Fanuc KAREL source: kd00051.KL

-- PROVISIONAL review KL for V940-1; original PC SHA256 1b8f119a18a5a4649315fc7f6d6ce60d3f234252100fceed115acb7b17a9f241
-- Incomplete behavior may be omitted. Consult companion uncertainty JSON. Do not deploy.
PROGRAM KD00051
%NOLOCKGROUP
VAR
  I : INTEGER
  J : INTEGER
  B : BOOLEAN
  R : REAL
  S : STRING[80]
-- UNRESOLVED_DECL P type=000101
BEGIN
  -- V9_ZERO_TABLE_METADATA_HINT layout=0001; no indexed target words; source/name/runtime held
  -- UNRESOLVED_PC offsets 5-30; opcodes 01,22,1C,2E,0A,82,0B
  -- UNRESOLVED_PC offsets 35-39; opcodes 7F
END KD00051
